// TIA Portal V21 export
// export: Created 2026-08-21T20:18:49.6575132Z, ExportSetting None, DisplayName Totally Integrated Automation Portal, DisplayVersion V21, DisplayName STEP 7 Professional, DisplayVersion V21, DisplayName STEP 7 Safety, DisplayVersion V21, DisplayName Tech WebApplication, DisplayVersion V21, DisplayName WinCC Basic/Comfort/Advanced, DisplayVersion V21, DisplayName WinCC Professional, DisplayVersion V21, DisplayName WinCC Unified, DisplayVersion V21
FUNCTION "AccuS_Liter" : Void   // FC12, FBD
{ S7_Optimized_Access := 'TRUE' }
// stored: SetENOAutomatically false
   VAR_TEMP
      State : "Service_States";
   END_VAR
   VAR_TEMP   // added for the SCL form of the ladder/FBD networks
      _w1 : Bool;
   END_VAR
BEGIN

REGION Network 1
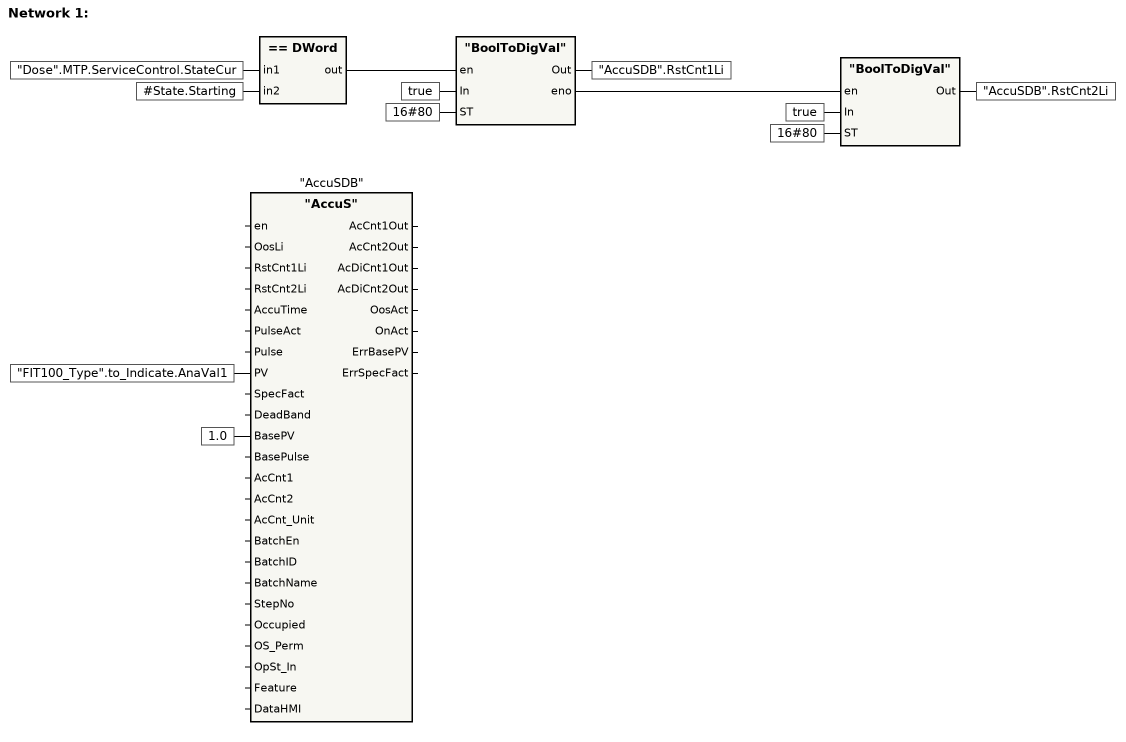
   "BoolToDigVal"(EN := "Dose".MTP.ServiceControl.StateCur = #State.Starting,
                  In := true,
                  ST := 16#80,
                  Out => "AccuSDB".RstCnt1Li,
                  ENO => #_w1);
   IF #_w1 THEN "BoolToDigVal"(In := true, ST := 16#80, Out => "AccuSDB".RstCnt2Li); END_IF;
   "AccuSDB"(PV := "FIT100_Type".to_Indicate.AnaVal1, BasePV := 1.0);   // "AccuS"
END_REGION
END_FUNCTION
